{attribute 'qualified_only'}
{attribute 'strict'}
{attribute 'to_string'}
TYPE E_Element_Process :
(
eNone := 0,
eDrain,
eWash_Recycle,
eWash_Detergent,
eWash_Water_1,
eWash_Sani,
eWash_Water_2,
eFill_Water,
eDissolving,
eConnectionToLine,
eDisconnection
);
END_TYPE

(* stored: Version 1.1.0.1, ProductVersion 3.1.4024.12
   DUT E_Element_Process: Id {b2ca1574-4be6-413a-9da5-e43d5cd3c451} *)
